{attribute 'qualified_only'}
{attribute 'strict'}
TYPE E_ASensor_State :
(
	Init := 0,
	Close,Open,Busy_Close,Busy_Open
);
END_TYPE

(* stored: Version 1.1.0.1, ProductVersion 3.1.4024.12
   EnumerationTextList E_ASensor_State: Id {5d6d33d6-06d6-437b-9a5e-01fafad11d77} *)
